Fanuc KAREL source: kt00605.KL

PROGRAM KT00605
%NOLOCKGROUP
VAR
I1:INTEGER;I2:INTEGER;OUT:REAL
BEGIN
--
--
I1=2
I2=3
I1=2
I2=3
OUT=((-I1))
END KT00605
